Fanuc KAREL source: ka00091.KL

-- PROVISIONAL review KL for V770-1; original PC SHA256 7f464457a1fc98e8995109bd03c6964fadafb260d5a98be57cea4992a5153dbf
-- Incomplete behavior may be omitted. Consult companion uncertainty JSON. Do not deploy.
PROGRAM KA00091
%NOLOCKGROUP
-- UNRESOLVED_DECL SRC type=000199
-- UNRESOLVED_DECL DST type=000106
BEGIN
  -- UNRESOLVED_PC offsets 5-25; opcodes 49,7E,4A
  -- UNRESOLVED_PC offsets 30-34; opcodes 7F
END KA00091
